FUNCTION_BLOCK VacuumCtrl (* Basic Function Block Type *)
  (* Standard: 61499-2 *)
  (* Version 0.0, 7/2/2026, Template *)
  PACKAGE Main;
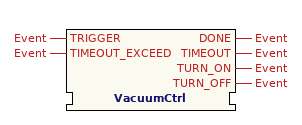
  EVENT_INPUT
    TRIGGER;
    TIMEOUT_EXCEED;
  END_EVENT
  EVENT_OUTPUT
    DONE;
    TIMEOUT;
    TURN_ON;
    TURN_OFF;
  END_EVENT
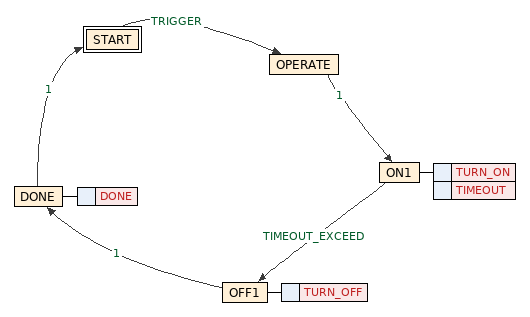
  EC_STATES
    START; (* Initial State *)
    OPERATE;
    ON1 : -> TURN_ON, -> TIMEOUT;
    OFF1 : -> TURN_OFF;
    DONE : -> DONE;
  END_STATES
  EC_TRANSITIONS
    START TO OPERATE := TRIGGER;
    OPERATE TO ON1 := 1;
    ON1 TO OFF1 := TIMEOUT_EXCEED;
    OFF1 TO DONE := 1;
    DONE TO START := 1;
  END_TRANSITIONS
  ALGORITHM INIT IN ST: (* Initialization algorithm *)
;
  END_ALGORITHM
  ALGORITHM REQ IN ST: (* Normally executed algorithm *)
;
  END_ALGORITHM
END_FUNCTION_BLOCK
